Fanuc KAREL source: KA00091.KL

PROGRAM KA00091
%NOLOCKGROUP
VAR
  SRC: JOINTPOS
  DST: XYZWPREXT
BEGIN
  DST = SRC
END KA00091
